(* IEC 61131-3 sources: daoli-st-library/DL_Device (part 41) *)

(* ---- FB_DL_OilLevelWatch.st ---- *)
(*
    FB_DL_OilLevelWatch —— 润滑 / 液压油油位连续监视（双阈值迟滞 + 确认延时 + NE107）
    ------------------------------------------------------------------
    组件名称  : FB_DL_OilLevelWatch
    分类      : DL_Device / LevelMonitoring
    前缀      : FB_DL_
    版本      : 1.0.0
    溯源      : 借鉴组织 —— T2-6 Rockwell AOI（矩阵行 166）：仅借鉴「设备级
                粗粒度监视 AOI」的公开功能形态（连续量监视 + 确认延时 +
                分级健康出口）；clean-room 声明 —— 零代码行复制，判据链 /
                迟滞口径 / 码位 100% 自有；非有限判据为 IEC 61131-3 标准语义
                （R79 双判）的道莅防御性实现。
    平台      : 纯 IEC 61131-3（TON / R_TRIG / LREAL 比较），CODESYS 3.5 /
                TwinCAT 3 / InoProShop / Machine Expert 通用
    作者      : 道莅代码库 · PLC编程专家（R72 构建轮 · 批 3 · 序号 9）
    ------------------------------------------------------------------
    功能说明  : 齿轮箱 / 液压单元油位巡检：欠油提前预警防干磨烧轴。
                单相监视（无顺序状态机 CASE，同族 FB_DL_AxisEncBatteryWatch
                口径家族一致）：
                ① 非有限液位闸：fLevelMm 非有限（NaN 自反判 + Inf 差值自反
                   判，R79）→ **直接故障锁存**（探头断线状态不明比欠油更
                   危险，R71 AxisEncBatteryWatch 口径家族一致），不等确认
                   延时；
                ② 组态域闸（R272 全枚举）：fLowWarnMm / fHystMm / fProbeMaxMm
                   非有限、fHystMm < 0（回差为负）、fLowWarnMm >= fProbeMaxMm
                   （阈值倒置）、fProbeMaxMm <= 0（量程非正）→ 组态锁存码
                   （根因优先归因，段 6 先于段 7）；
                ③ 双阈值迟滞判定：未预警相以进入线判（fLevelMm < fLowWarnMm），
                   已预警相以退出线判（fLevelMm >= fLowWarnMm + fHystMm），
                   防临界抖振；
                ④ TON 连续确认（断输入口径：液位回升出迟滞带 IN 即 FALSE，
                   计时清零重计）→ 预警锁存；
                ⑤ NE107 健康出口：欠油确认 → eMaintenanceReq；非有限 /
                   组态故障 → eFailure；正常 → eOk；失能 → eCheckFunction。
                锁存解除口径（R321 电平式声明）：bReset 上升沿为**唯一人工
                解除**，液位恢复越退出线为**条件恢复自动降级**双路——两路
                并存写死，禁恢复沿作唯一解除载体。预警锁存后自动降级判据 =
                液位 >= 退出线（迟滞带内保持预警，出带即自动解除）。
                满油探头饱和：fLevelMm > fProbeMaxMm → 信息级（满油合法
                工况，不拦截照判——判定方向与液位单调性一致，无危险侧偏差）。
                失能语义（R191 声明）：bEn = FALSE → bLowWarn / bError /
                nErrCode 出口清零、eHealth = eCheckFunction；_bFault /
                _bWarnLatch 锁存位**不被失能清除**（失能是操作态不是复位），
                须 bReset 上升沿解除——两语义分离。
    错误码    : 16#0003_0740 液位非有限（探头断线 / ADC 故障），直接锁存不等
                            确认延时 —— 故障级
                16#0003_0741 组态非法（阈值倒置 / 回差为负 / 阈值或量程非有限 /
                            量程非正 / 预警线不低量程上界），锁存至复位沿
                            —— 故障级
                16#0003_0742 液位越探头量程上界（探头饱和，满油合法工况）
                            —— 信息级，不置 bError（R45）
                加码反证句（R90）：0740（探头）与 0741（组态）成因互斥且调用
                方可自证（接线 vs 组态表），eHealth 出口同为 eFailure 但码位
                分流维修动作，输出组合不可互换观测，故各立一码；0742 由
                「液位在迟滞带上方 + 码位非零」唯一观测（正常满油不带码），
                不与既有输出组合重复。
    码位总账  : 16#0003_0740 用 ｜ 16#0003_0741 用 ｜ 16#0003_0742 用
    状态机    : N/A —— 单相监视，无顺序状态机，无自有 ENUM / CASE 可写；
                确认计时由 TON 实例自持（定时器状态而非顺序状态）；
                健康出口复用既有枚举 E_DL_Ne107Status（只引用）
    边界与披露: 一 TON（tonConfirm）与 R_TRIG（rtReset）每拍**无条件调用**
                   （规则 ⑦），IN 为段 7 计算出的显式条件；
                二 零全局变量、零 VAR_EXTERNAL、零物理地址；
                三 归属 Ownership：E_DL_Ne107Status 归属 I_DL_DeviceHealth.st
                   （全库唯一定义，R264），本件只引用不重声明；
                四 输入非有限 / 组态非法 → 直接锁存（不走迟滞判定集合，安全
                   侧赋值不引用本闸判定内的量，防自证循环，R127）；
                五 输出量纲：fLevelMm / fLowWarnMm / fHystMm / fProbeMaxMm 均
                   [mm]，本件不换算单位；
                六 分工互引：FB_DL_SiloLevelInterlock（料仓联锁）、
                   FB_DL_LevelSwitchVib（开关量检测）、FB_DL_HydrostaticLevelComp
                   （静压补偿换算）——本件只做模拟量油位趋势监视，不做联锁
                   与换算；
                七 依赖声明：仅 Standard.library（TON / R_TRIG / ABS），零
                   厂商方言。
    验收向量  : V1 液位 80 mm、预警线 100 mm、确认 2 s → 2 s 后 bLowWarn；
                V2 液位回升 130 mm（退出线 100 + 20）→ 自动降级解除；
                V3 液位回升 110 mm（迟滞带内）→ 预警保持（迟滞自证）；
                V4 fLevelMm = NaN → 0740 立即锁存（不等 2 s）；V5 fHystMm
                = −1 → 0741 锁存；V6 fLevelMm = 520（量程 500）→ 0742
                信息级照判；V7 bReset 上升沿 → 清锁存；V8 失能 → 出口清零、
                锁存保留。
                算法已证（脚本）：未跑 ｜ 编译器已证（三平台）：未跑
    修订记录  : 2026-11-23 v1.0.0 首次入库（R72 构建轮 · 批 3 · 序号 9）
*)
FUNCTION_BLOCK FB_DL_OilLevelWatch
VAR_INPUT
    fLevelMm    : LREAL;                   (* 油位连续值（引脚注入），[mm]，非有限即探头故障 / the oil level continuous value in mm *)
    fLowWarnMm  : LREAL := 100.0;          (* 低油位预警阈值（迟滞进入线），[mm] / the low oil warn threshold, the hysteresis enter line *)
    fHystMm     : LREAL := 20.0;           (* 迟滞回差（退出线 = 预警线 + 回差），[mm]，禁负 / the hysteresis band in mm, the exit line is warn plus band *)
    fProbeMaxMm : LREAL := 500.0;          (* 探头量程上界（饱和信息级判据），[mm]，禁非正 / the probe range upper bound in mm *)
    tConfirm    : TIME := T#2S;            (* 欠油确认延时，[ms] / the low oil confirmation delay *)
    bEn         : BOOL := TRUE;            (* 使能，[标志]，FALSE 出口清零、锁存保留 / the enable, FALSE clears the outlets, the latch kept *)
    bReset      : BOOL := FALSE;           (* 故障 / 预警复位，[标志]，上升沿唯一人工解除 / the reset, its rising edge is the only manual release *)
END_VAR
VAR_OUTPUT
    bLowWarn  : BOOL := FALSE;             (* 低油位预警锁存位（确认成立且未解除）[标志] / the low oil warn latched flag *)
    eHealth   : E_DL_Ne107Status;          (* NE107 健康出口（欠油 → eMaintenanceReq，故障 → eFailure）/ the NE 107 health outlet *)
    bValid    : BOOL := FALSE;             (* 出口可用标志，失能或锁存故障为 FALSE / the outlets usable *)
    bError    : BOOL := FALSE;             (* 故障标志，存在锁存故障时 TRUE / the fault flag *)
    nErrCode  : UDINT := 16#0000_0000;     (* 错误码，0 = 正常，锁存回放（R187）/ the error id, replayed from the latch *)
END_VAR
VAR
    _rtReset    : R_TRIG;                  (* 复位上升沿实例（无条件调用）/ the reset rising edge instance *)
    _tonConfirm : TON;                     (* 欠油确认延时实例（无条件调用）/ the low oil confirmation timer *)
    _bFault     : BOOL := FALSE;           (* 故障锁存副本（探头 / 组态），仅复位沿解除 / the internal fault latch copy *)
    _nCodeLatch : UDINT := 0;              (* 锁存成因码，故障期回放 / the latched cause code *)
    _bWarnLatch : BOOL := FALSE;           (* 预警锁存副本（自动降级或复位沿解除）/ the warn latch copy *)
    _bCfgBad    : BOOL := FALSE;           (* 组态非法标志（逐拍重算，仅用于首次锁存）/ the config fault flag *)
    _bInBad     : BOOL := FALSE;           (* 液位非有限标志（逐拍重算）/ the input fault flag *)
    _bOutDom    : BOOL := FALSE;           (* 液位越量程上界标志（逐拍重算，信息级）/ the probe saturation flag *)
    _bRun       : BOOL := FALSE;           (* 运行许可 = 使能 且 无锁存故障 / the run permit *)
    _bLowCond   : BOOL := FALSE;           (* 欠油迟滞判定条件（含自保持，送 TON）/ the low oil hysteresis condition *)
END_VAR
VAR CONSTANT
    DL_OLW_CODE_PROBE : UDINT := 16#0003_0740; (* 液位非有限锁存码 [码] / the probe fault code *)
    DL_OLW_CODE_CFG   : UDINT := 16#0003_0741; (* 组态非法锁存码 [码] / the configuration fault code *)
    DL_OLW_CODE_SAT   : UDINT := 16#0003_0742; (* 探头饱和信息码 [码] / the probe saturation info code *)
    DL_OLW_ZERO       : UDINT := 0;            (* 无符号零哨兵 [码] / the unsigned zero sentinel *)
    DL_OLW_FZERO      : LREAL := 0.0;          (* 浮点零哨兵 [mm] / the float zero sentinel *)
END_VAR

// 段 1｜出口预置（统一出口预置，R256）/ segment 1, preset every outlet
bLowWarn := FALSE;                         // 预警出口预清零（映射段回填）/ preset the warn outlet false
eHealth  := E_DL_Ne107Status.eUnknown;     // 健康出口预置未知（首拍语义）/ preset the health outlet unknown
bValid   := FALSE;                         // 可用标志预清零 / preset the usable flag false
bError   := FALSE;                         // 故障标志预清零 / preset the fault flag false
nErrCode := DL_OLW_ZERO;                   // 码位预置无错 / preset the code zero
_bLowCond := FALSE;                        // 迟滞条件预清零 / preset the condition false

// 段 2｜复位沿无条件调用（规则 ⑦）/ segment 2, the unconditional reset edge refresh
_rtReset(CLK := bReset);                   // 每拍无条件刷新 / refreshed every scan

// 段 3｜锁存解除：复位沿唯一人工解除（作用域：清双锁存 + 清码，R311 声明）/ segment 3, the manual release edge
IF _rtReset.Q THEN                         // 复位上升沿 / the reset rising edge
    _bFault := FALSE;                      // 清故障锁存（恒可达，R152 自证）/ clear the fault latch
    _bWarnLatch := FALSE;                  // 清预警锁存 / clear the warn latch
    _nCodeLatch := DL_OLW_ZERO;            // 清锁存码（可到达清除边）/ clear the latched code
END_IF

// 段 4｜组态域闸（R272 全枚举：fLowWarnMm / fHystMm / fProbeMaxMm 三引脚）/ segment 4, the configuration guard
_bCfgBad := (fLowWarnMm <> fLowWarnMm) OR ((fLowWarnMm - fLowWarnMm) <> DL_OLW_FZERO) // 预警线非有限 / the warn line non finite
         OR (fHystMm <> fHystMm) OR ((fHystMm - fHystMm) <> DL_OLW_FZERO)              // 回差非有限 / the hysteresis non finite
         OR (fProbeMaxMm <> fProbeMaxMm) OR ((fProbeMaxMm - fProbeMaxMm) <> DL_OLW_FZERO) // 量程非有限 / the range non finite
         OR (fHystMm < DL_OLW_FZERO)                                                   // 回差为负 / a negative hysteresis
         OR (fLowWarnMm >= fProbeMaxMm)                                                // 阈值倒置（预警线不低于量程上界）/ the threshold inversion
         OR (fProbeMaxMm <= DL_OLW_FZERO);                                             // 量程非正 / a non positive range

// 段 5｜输入守卫：液位非有限即危险（状态不明 > 欠油，直接锁存不等延时）/ segment 5, the input guard
_bInBad := (fLevelMm <> fLevelMm) OR ((fLevelMm - fLevelMm) <> DL_OLW_FZERO); // 液位非有限（R79 双判）/ the level non finite
_bOutDom := (fLevelMm > fProbeMaxMm);      // 液位越量程上界（探头饱和，信息级）/ the level over the range

// 段 6｜首次成因锁存（故障期内不重推断，回放锁存码，R189；组态根因优先）/ segment 6, the first cause latch
IF NOT _bFault THEN                        // 未锁存才登记 / register only while not latched
    IF _bCfgBad THEN                       // 组态非法（根因优先归因）/ the config fault first
        _bFault := TRUE;                   // 置锁存 / latch
        _nCodeLatch := DL_OLW_CODE_CFG;    // 登记组态码 / register the config code
    ELSIF _bInBad THEN                     // 液位非有限（不等确认延时）/ the probe fault, no delay
        _bFault := TRUE;                   // 置锁存 / latch
        _nCodeLatch := DL_OLW_CODE_PROBE;  // 登记探头码 / register the probe code
    END_IF
END_IF

// 段 7｜运行许可与迟滞条件（分支内不调用任何定时器）/ segment 7, the run permit and the hysteresis condition
_bRun := bEn AND (NOT _bFault);            // 使能且无锁存故障 / enabled and not latched
IF _bRun THEN                              // 运行许可成立 / the run permit holds
    IF _bWarnLatch THEN                    // 已预警相：以退出线判（迟滞防抖振）/ the latched phase, the exit line
        _bLowCond := fLevelMm < (fLowWarnMm + fHystMm); // 迟滞带内保持预警 / hold inside the band
    ELSE                                   // 未预警相：以进入线判 / the unlatched phase, the enter line
        _bLowCond := fLevelMm < fLowWarnMm; // 破进入线 / under the enter line
    END_IF
    IF _bLowCond AND _tonConfirm.Q THEN    // 破线经确认延时 / the condition confirmed
        _bWarnLatch := TRUE;               // 预警锁存 / latch the warn
    END_IF
    IF _bWarnLatch AND (NOT _bLowCond) THEN // 条件恢复自动降级（电平式双路之二，R321 声明；复位沿为人工路）/ the automatic level release
        _bWarnLatch := FALSE;              // 出迟滞带即自动解除（同拍生效）/ release over the exit line
    END_IF
ELSE                                       // 失能或锁存故障 / disabled or latched
    _bLowCond := FALSE;                    // 条件清零（TON 随之复位）/ clear the condition
END_IF

// 段 8｜确认定时器无条件调用（IN 为段 7 显式条件；断输入口径：出线即断计）/ segment 8, the unconditional confirmation timer
_tonConfirm(IN := _bRun AND _bLowCond, PT := tConfirm); // 欠油确认计时 / the confirmation timer

// 段 9｜出口映射（名实双出口同源，R191）/ segment 9, the outlet mapping
IF _bRun THEN                              // 运行许可成立 / the run permit holds
    bLowWarn := _bWarnLatch;               // 预警出口与锁存同源 / the warn outlet shares the latch
    bValid := TRUE;                        // 出口可用 / the outlets usable
    IF _bWarnLatch THEN                    // 预警确认成立 / the warn confirmed
        nErrCode := DL_OLW_ZERO;           // 预警本身不发码（欠油是正常工况分支非缺陷）/ the warn carries no code
        eHealth := E_DL_Ne107Status.eMaintenanceReq; // 欠油 → 需要维护 / maintenance required
    ELSE                                   // 无预警 / no warn
        eHealth := E_DL_Ne107Status.eOk;   // 正常 / ok
    END_IF
    IF _bOutDom AND (NOT _bWarnLatch) THEN // 运行中探头饱和且无更高优先级出口 / the saturation info
        nErrCode := DL_OLW_CODE_SAT;       // 信息级：探头饱和满油（不置 bError，R45）/ info level: the probe saturation
    END_IF
ELSIF (NOT bEn) THEN                       // 失能相（操作态优先于故障归因，同族口径）/ the disabled phase
    bLowWarn := FALSE;                     // 出口清零（锁存保留）/ the outlet cleared, the latch kept
    bError := FALSE;                       // 失能不是故障 / a disabled block is not a fault
    nErrCode := DL_OLW_ZERO;               // 失能不发码 / no code while disabled
    eHealth := E_DL_Ne107Status.eCheckFunction; // 失能 → 功能检查 / function check
ELSE                                       // 锁存故障相（失能优先级之上）/ the latched fault phase
    bLowWarn := FALSE;                     // 故障相预警出口清零（归并故障出口）/ the warn outlet cleared
    bError := TRUE;                        // 故障标志置位 / raise the fault flag
    nErrCode := _nCodeLatch;               // 回放锁存码 / replay the latched code
    eHealth := E_DL_Ne107Status.eFailure;  // 故障 → 失效（信号不可信）/ failure
END_IF
END_FUNCTION_BLOCK

(* ---- FB_DL_PressureReliefMonitor.st ---- *)
(*==============================================================================
 * 组件名称 (Component)  : FB_DL_PressureReliefMonitor
 * 溯源说明 (Provenance): 道莅 clean-room 防御性实现（IEC 61131-3 纯净实现，闭源文档仅借语义，零代码行）
 * 所属子库 (Sublibrary) : DL_Device / SafetyMonitor
 * 当前版本 (Version)    : 1.0.0
 * 兼容性   (Platform)   : CODESYS 3.5 / TwinCAT 3 / 汇川 InoProShop / 施耐德
 *                         Machine Expert；纯 IEC 61131-3（第 3 版），仅用
 *                         Standard.library 的 TON / ABS / MAX
 * 组件分类 (Category)   : 功能块（FUNCTION_BLOCK）· 安全阀起跳/回座监视与台账
 * 功能一句话 (Summary)  : 用阀前/阀后压力判安全阀是否起跳，累计动作次数与累计
 *                         开启时长，给出本次起跳峰值压力与 NE107 健康分级。
 *
 * 本件存在的意义 (Why this unit exists)
 *   过程安全台账要求「安全阀一年动作了几次、累计开启多久」——这是法检项。
 *   库内 AlarmManager 数的是报警不是阀门动作，PortDiag 系列数的是通讯事件，
 *   没有任何件维护这张台账。同时「阀前持续超整定而阀后不同步升高」是
 *   安全阀不泄放的典型特征，属于必须报出来的失效形态。
 *
 * 台账纪律 (Ledger discipline)
 *   ① 起跳判据必须用**回座比做迟滞**（fUpPressure < fSetPressure × fBlowdown），
 *      硬阈值会让压力在整定点附近抖动并反复计数——这是台账失真的头号原因；
 *   ② 单次起跳时长 < tMinLift 不计入 nLiftCount（信息 0175）：工艺压力波动
 *      引起的瞬时顶开不构成「动作」，但仍计入累计开启时长之外的判定之外，
 *      两者口径不同，头注释写死；
 *   ③ 计数与累计时长累加前判上界，饱和不回绕（R35）；TIME 溢出用比较式
 *      预判（R54），比较表达式内不出现加乘运算符；
 *   ④ **失能不清台账**：计数、累计时长、峰值一律保持；若失能发生在起跳期间，
 *      以失能拍作为该次起跳的结束拍如实入账，绝不丢一次真实动作。
 *
 * 健康映射（写死在此，不散落实现体）
 *   参数非法 / 输入非有限                        → eFailure
 *   起跳中且阀后压力 > 整定 × DL_DN_FAIL_RATIO    → eFailure（疑似不泄放）
 *   nLiftCount >= uMaintLimit                    → eMaintenanceReq
 *   其余（有判定能力）                            → eOk
 *   未使能（无判定能力）                          → eUnknown
 *   DL_DN_FAIL_RATIO = 0.5 为件内经验阈值：安全阀正常起跳时阀后应接近大气，
 *   若阀后压力仍高于整定的一半，说明介质没有真正排出去（下游堵塞或阀瓣卡滞）。
 *
 * 边界安全 (Boundary)
 *   - fSetPressure <= 0 或 fBlowdown 不在 (0, 1) 或非有限 → 故障 033F、bValid = FALSE，
 *     **台账保持不动**（参数错了不等于阀门没动作过）；
 *   - 任一压力非有限 → 故障 0340，**保持 bLifted 与计数不变**（坏值不得伪造动作）；
 *   - bError 的每一个置位源都能在 eErr 找到对应码（R45 纪律）；
 *   - CASE 落 ELSE 置 0341 兜底并回 eFault；
 *   - 本件无复位引脚：台账只能靠 FB 实例重建清零（法检台账不允许被误复位，
 *     这是刻意设计，已留档）。
 *
 * 错误码    : 16#0003_0174 起跳事件已记录（动作次数 +1，累计时长继续累加）——信息级
 *             16#0003_0175 单次起跳时长低于 tMinLift，按工艺波动滤除不计入台账——信息级
 *             16#0003_033F 整定压力或回座比非法——故障级，bValid = FALSE
 *             16#0003_0340 压力输入非有限，保持台账与判定不变——故障级，坏值不得伪造动作
 *             16#0003_0341 状态机落 ELSE 兜底（非法状态）——故障级，回 eIdle 并保持台账
 * 码位总账  : 16#0003_0174 用 / 16#0003_0175 用 ｜ 16#0003_033F 用 / 16#0003_0340 用 / 16#0003_0341 用
 * 状态机    : E_DL_ReliefState（eIdle / eLifted / eReseat / eFault），CASE 含 ELSE 兜底，
 *             ELSE 置 16#0003_0341 并回 eFault；失能回 eIdle 但台账保持
 * 采样约定  : 每任务周期调用一次；时长按滚动时钟差累加（上拍快照，R45②）
 * 依赖说明  : 仅 Standard.library；健康出口引用 E_DL_Ne107Status（属主 I_DL_DeviceHealth，
 *             **引用不重声明**，R70③）
 * 验收向量  : V1 压力从 8 缓升到 10.5 bar 持续 200 ms → eLifted，bLifted = TRUE，
 *                fPeakPressure 跟随峰值；压力回落到 8.9（< 10×0.90 = 9.0）→ eReseat，
 *                时长 ≥ 500 ms 时 nLiftCount + 1 且 eErr = 0174，eHealth 随计数升级
 *             V2 起跳仅 300 ms（< tMinLift 500 ms）→ nLiftCount 不变，eErr = 0175（滤除主向量）
 *             V3 起跳中阀后压力 6 bar（> 10×0.5）→ eHealth = eFailure（不泄放主向量）
 *             V4 fBlowdown = 1.2 → 033F，bValid = FALSE，nLiftCount 与 tOpenTotal 保持
 *             V5 fUpPressure = NaN → 0340，bLifted 与计数保持（坏值不伪造动作主向量）
 *             V6 压力在 9.98~10.02 之间抖动 → 不重复计数（回座迟滞主向量）
 *             V7 bEnable 落于起跳中 → eIdle，本次时长如实入账，计数不清零
 * 红线自检  : 全局变量声明零使用 / 外部变量访问零使用 / 物理地址零使用 ｜ 纯 IEC 61131-3 ｜ 无除法
 *             浮点只用大小与容差比较 ｜ 无循环 ｜ 全变量双语同行注释 ｜ ENUM + CASE
 *             含 ELSE ｜ TON 在主体前部无条件刷新 ｜ TIME 溢出比较式预判 ｜
 *             阈值常量化，无魔法数
 * 修订历史  : 2026-11-16  v1.0.0  首版入库（R22 · 批 2 · 设备安全台账）
 *============================================================================*)

(*-----------------------------------------------------------------------------
 * 枚举: E_DL_ReliefState（归属本功能块，同文件发布，全库唯一定义）
 * 含义: 安全阀监视的工作相位。0 起步长 10。
 * 注意: 健康出口类型 E_DL_Ne107Status 属主为 I_DL_DeviceHealth（DL_Device 契约件），
 *       本件只引用、不重声明（R70③ 全库唯一定义）。
 *-----------------------------------------------------------------------------*)
TYPE E_DL_ReliefState :
(
    eIdle   := 0,      // 待机：未起跳，等待起跳确认 / Idle, waiting for a confirmed lift
    eLifted := 10,     // 起跳中：阀前高于整定，正在累计时长 / Lifted, upstream above the set pressure
    eReseat := 20,     // 回座：单拍入账相，随后回待机 / Reseat, one scan to book the event
    eFault  := 99      // 故障：参数非法或输入非有限 / Fault, illegal parameter or non-finite input
);
END_TYPE

FUNCTION_BLOCK FB_DL_PressureReliefMonitor
VAR_INPUT
    fUpPressure  : REAL;                       // 阀前压力 [bar g] / upstream pressure [bar g]
    fDnPressure  : REAL;                       // 阀后压力 [bar g] / downstream pressure [bar g]
    fSetPressure : REAL := 10.0;               // 整定压力 [bar g]，须 > 0 / set pressure [bar g], must be > 0
    fBlowdown    : REAL := 0.90;               // 回座压力比 [倍]，须在 0~1 之间 / reseat ratio [ratio], must lie inside zero and one
    tConfirm     : TIME := T#200MS;            // 起跳确认时间 [ms] / lift confirm time [ms]
    tMinLift     : TIME := T#500MS;            // 最短起跳时长 [ms]，低于此按波动滤除 / minimum lift duration [ms], shorter ones are filtered
    uMaintLimit  : UINT := 50;                 // 动作次数维护门限 [次] / maintenance count threshold [count]
    bEnable      : BOOL;                       // 使能（失能不清台账） / enable, the ledger survives a disable
END_VAR
VAR_OUTPUT
    bLifted      : BOOL;                       // 当前处于起跳状态 / currently lifted
    nLiftCount   : UDINT;                      // 累计动作次数 [次] / accumulated lift count [count]
    tOpenTotal   : TIME;                       // 累计开启时长 [ms] / accumulated open time [ms]
    fPeakPressure : REAL;                      // 本次起跳峰值压力 [bar g] / peak upstream pressure of the current lift [bar g]
    eHealth      : E_DL_Ne107Status;           // NE107 健康分级（引用唯一属主） / NE107 health status, referenced from its owner
    eErr         : UDINT;                      // 错误码，0 表示无错 / error code, 0 means no error
    bError       : BOOL;                       // 故障级标志，仅故障级错误置位 / fault-class flag, set only on fault-level codes
    bValid       : BOOL;                       // 输出可用标志 / outputs usable flag
END_VAR
VAR
    fbConfirm    : TON;                        // 起跳确认计时，段 5 无条件刷新 [ms] / lift confirm timer
    fbElapsed    : TON;                        // 滚动时钟，段 5 无条件刷新 [ms] / rolling elapsed clock
    _eState      : E_DL_ReliefState := E_DL_ReliefState.eIdle; // 当前相位 / current phase
    _bInit       : BOOL := FALSE;              // 首扫标志，初值 FALSE 取非判定 / first-scan flag, tested negated
    _bParamBad   : BOOL;                       // 参数非法标志 / illegal parameter flag
    _bFiniteBad  : BOOL;                       // 输入非有限标志 / non-finite input flag
    _bIllegal    : BOOL;                       // 非法状态标志 / illegal state flag
    _bAbove      : BOOL;                       // 阀前高于整定（确认条件） / upstream above the set pressure
    _bReseatNow  : BOOL;                       // 回座判据成立 / reseat criterion satisfied
    _bConfBreak  : BOOL;                       // 确认计时器断输入一拍 / confirm timer one-scan break
    _bElapsedBreak : BOOL;                     // 滚动时钟断输入一拍 / rolling clock one-scan break
    _bNoRelief   : BOOL;                       // 疑似不泄放标志 / suspected no-relief flag
    _bBooked     : BOOL;                       // 本拍已入账标志 / booked this scan flag
    _bReseatPulse : BOOL;                      // 回座单拍脉冲（入账触发） / reseat one-scan pulse, triggers the booking
    _bLiftedPrev : BOOL;                       // 本拍进入时的起跳相快照（R38 镜像量） / lifted snapshot taken before the transitions
    _tConfirmUse : TIME := T#200MS;            // 生效确认时间 [ms]，已钳位 / effective confirm time, clamped
    _tMinLiftUse : TIME := T#500MS;            // 生效最短起跳时长 [ms]，已钳位 / effective minimum lift, clamped
    _tEtPrev     : TIME;                       // 滚动时钟上拍快照 [ms] / previous scan snapshot of the clock
    _tDelta      : TIME;                       // 本拍时长增量 [ms] / elapsed increment of this scan
    _tLiftDur    : TIME;                       // 本次起跳已持续时长 [ms] / duration of the current lift [ms]
    _tTotalAcc   : TIME;                       // 累计开启时长保持量 [ms] / held accumulated open time [ms]
    _uCountAcc   : UDINT;                      // 累计动作次数保持量 [次] / held lift count [count]
    _fPeakAcc    : REAL;                       // 本次起跳峰值保持量 [bar g] / held peak pressure of the current lift [bar g]
    _fPeakTot    : REAL;                       // 历史峰值（供 HMI 参考） [bar g] / historical peak pressure [bar g]
END_VAR
VAR CONSTANT
    DL_VAL_LIM   : REAL := 1.0E6;              // 有限性判定的绝对值上限 [bar g] / finiteness ceiling [bar g]
    DL_SET_MIN   : REAL := 0.0;                // 整定压力下限 [bar g]，须严格大于 / set pressure floor, strictly greater
    DL_BLOW_MIN  : REAL := 0.0;                // 回座比下限 [倍]，须严格大于 / reseat ratio floor, strictly greater
    DL_BLOW_MAX  : REAL := 1.0;                // 回座比上限 [倍]，须严格小于 / reseat ratio ceiling, strictly less
    DL_DN_FAIL_RATIO : REAL := 0.5;            // 阀后不泄放判据比 [倍]，件内经验阈值 / no-relief ratio, an empirical in-unit threshold
    DL_CONF_MAX_MS : DINT := 60000;            // 确认时间上限 [ms] / confirm time ceiling [ms]
    DL_MINLIFT_MAX_MS : DINT := 3600000;       // 最短起跳时长上限 [ms]，一小时 / minimum lift ceiling, one hour
    DL_TIME_ZERO : TIME := T#0MS;              // 时间零值基准 [ms] / time zero reference
    DL_ROLL      : TIME := T#1H;               // 滚动时钟周期 [ms]，到顶重启防 ET 停滞 / rolling clock period, restarted at the top
    DL_TOTAL_MAX : TIME := T#24H;              // 累计时长饱和上界 [ms] 上限值：判溢出用 / accumulation ceiling, used by the overflow test
    DL_TIME_SAT  : TIME := T#24H;              // 累计时长饱和输出值 [ms] / accumulation saturation value
    DL_CNT_MAX   : UDINT := 16#FFFF_FFFF;      // 计数饱和上界 [次]，不回绕 / counter saturation ceiling, never wraps
END_VAR

(*------------------------------------------------------------------------------
 * 段 1｜每拍预置（台账保持量不预置；输出在段 9 单点写入）
 *      Per-scan presets, the ledger values are never cleared here
 *-----------------------------------------------------------------------------*)
eErr         := 16#0000_0000;                  // 错误码每拍重算 / error code recomputed every scan
bError       := FALSE;                         // 故障标志每拍重算 / fault flag recomputed every scan
bValid       := FALSE;                         // 可用标志每拍重算 / usable flag recomputed every scan
_bParamBad   := FALSE;                         // 参数非法标志预清零 / parameter flag pre-cleared
_bFiniteBad  := FALSE;                         // 非有限标志预清零 / non-finite flag pre-cleared
_bIllegal    := FALSE;                         // 非法状态标志预清零 / illegal state flag pre-cleared
_bAbove      := FALSE;                         // 超整定条件预置 FALSE / above-set condition preset FALSE
_bReseatNow  := FALSE;                         // 回座判据预置 FALSE / reseat criterion preset FALSE
_bNoRelief   := FALSE;                         // 不泄放标志预置 FALSE / no-relief preset FALSE
_bBooked     := FALSE;                         // 入账标志预置 FALSE / booked flag preset FALSE
_bReseatPulse := FALSE;                        // 回座脉冲预置 FALSE / reseat pulse preset FALSE
_bLiftedPrev := FALSE;                         // 起跳快照预置 FALSE / lifted snapshot preset FALSE

(*------------------------------------------------------------------------------
 * 段 2｜首扫初始化（台账全部从零起，峰值从当前阀前压力起）
 *      First-scan initialisation, the ledger starts at zero
 *-----------------------------------------------------------------------------*)
IF NOT _bInit THEN
    _eState     := E_DL_ReliefState.eIdle;     // 相位待机 / phase idle
    _uCountAcc  := 0;                          // 动作次数清零 [次] / lift count cleared
    _tTotalAcc  := DL_TIME_ZERO;               // 累计时长清零 [ms] / accumulated time cleared
    _tLiftDur   := DL_TIME_ZERO;               // 本次时长清零 [ms] / current lift duration cleared
    _tEtPrev    := DL_TIME_ZERO;               // 时钟快照清零 [ms] / clock snapshot cleared
    _fPeakAcc   := 0.0;                        // 本次峰值清零 [bar g] / current peak cleared
    _fPeakTot   := 0.0;                        // 历史峰值清零 [bar g] / historical peak cleared
    _bConfBreak := TRUE;                       // 确认计时从零开始 / confirm timer starts from zero
    _bElapsedBreak := TRUE;                    // 滚动时钟从零开始 / rolling clock starts from zero
    _bInit      := TRUE;                       // 首扫只做一次 / the first scan runs once
END_IF

(*------------------------------------------------------------------------------
 * 段 3｜参数闸门（整定压力与回座比；非法只降可用性，台账一律保持）
 *      Parameter gate, an illegal parameter lowers usability but never touches the ledger
 *-----------------------------------------------------------------------------*)
IF (fSetPressure <> fSetPressure) OR (ABS(fSetPressure) > DL_VAL_LIM) OR (fSetPressure <= DL_SET_MIN) THEN
    _bParamBad := TRUE;                        // 整定压力非法 / set pressure illegal
END_IF
IF (fBlowdown <> fBlowdown) OR (fBlowdown <= DL_BLOW_MIN) OR (fBlowdown >= DL_BLOW_MAX) THEN
    _bParamBad := TRUE;                        // 回座比非法（须严格在 0~1 之间） / reseat ratio illegal
END_IF

(*------------------------------------------------------------------------------
 * 段 4｜压力输入有限性（区间判据同时拦 NaN 与 ±Inf）
 *      Pressure finiteness, the interval test catches NaN and infinity
 *-----------------------------------------------------------------------------*)
IF (fUpPressure < -DL_VAL_LIM) OR (fUpPressure > DL_VAL_LIM) THEN
    _bFiniteBad := TRUE;                       // 阀前压力非有限 / upstream pressure non-finite
END_IF
IF (fDnPressure < -DL_VAL_LIM) OR (fDnPressure > DL_VAL_LIM) THEN
    _bFiniteBad := TRUE;                       // 阀后压力非有限 / downstream pressure non-finite
END_IF

(*------------------------------------------------------------------------------
 * 段 5｜计时器无条件刷新（R40）+ 本拍时长增量（R45② 上拍快照）
 *      Timers refreshed unconditionally, the elapsed increment uses a previous-scan snapshot
 *-----------------------------------------------------------------------------*)
_tConfirmUse := tConfirm;                      // 确认时间直取引脚 [ms] / confirm time from the pin
IF TIME_TO_DINT(_tConfirmUse) > DL_CONF_MAX_MS THEN
    _tConfirmUse := DINT_TO_TIME(DL_CONF_MAX_MS); // 超上限钳位（无专用码位，R90 不新开码） / clamped
END_IF
IF TIME_TO_DINT(_tConfirmUse) < 0 THEN
    _tConfirmUse := DL_TIME_ZERO;              // 负时间结构性不可达，兜底为 0 / structurally unreachable fallback
END_IF

_tMinLiftUse := tMinLift;                      // 最短起跳时长直取引脚 [ms] / minimum lift from the pin
IF TIME_TO_DINT(_tMinLiftUse) > DL_MINLIFT_MAX_MS THEN
    _tMinLiftUse := DINT_TO_TIME(DL_MINLIFT_MAX_MS); // 超上限钳位 / clamped
END_IF
IF TIME_TO_DINT(_tMinLiftUse) < 0 THEN
    _tMinLiftUse := DL_TIME_ZERO;              // 负时间兜底为 0 / fallback to zero
END_IF

IF NOT _bFiniteBad THEN
    _bAbove := (fUpPressure > fSetPressure);   // 超整定判据 [布尔] / above-set test
    IF NOT _bParamBad THEN
        _bReseatNow := (fUpPressure < (fSetPressure * fBlowdown)); // 回座判据：低于整定×回座比 / reseat test
    END_IF
    _bNoRelief := (fDnPressure > (fSetPressure * DL_DN_FAIL_RATIO)); // 阀后未降：疑似不泄放 / downstream not relieved
END_IF

fbConfirm(IN := _bAbove AND (NOT _bConfBreak), PT := _tConfirmUse); // 起跳确认计时
_bConfBreak := FALSE;                          // 断输入拍在调用后自清 / break self-cleared after the call

fbElapsed(IN := (NOT _bElapsedBreak), PT := DL_ROLL); // 滚动时钟无条件刷新
_bElapsedBreak := FALSE;                       // 断输入拍在调用后自清 / break self-cleared
_tDelta := fbElapsed.ET - _tEtPrev;            // 本拍增量 = 当前 ET − 上拍快照 / increment from the snapshot
IF TIME_TO_DINT(_tDelta) < 0 THEN
    _tDelta := DL_TIME_ZERO;                   // 时钟重启拍：增量按 0 处理，绝不倒扣 / restart scan counts as zero
END_IF
_tEtPrev := fbElapsed.ET;                      // 快照在本拍末更新（唯一写入点） / snapshot updated once
IF fbElapsed.Q THEN
    _bElapsedBreak := TRUE;                    // 到顶重启：下一拍 ET 归零 / restart so the next scan starts from zero
    _tEtPrev := DL_TIME_ZERO;                  // 重启后快照同步归零 / the snapshot follows the restart
END_IF

(* 起跳相快照在迁移之前采集（R38）：迁移拍也要把本拍时长增量算进本次起跳 *)
(* The lifted snapshot is taken before the transitions so the final scan still counts *)
_bLiftedPrev := (_eState = E_DL_ReliefState.eLifted);

(*------------------------------------------------------------------------------
 * 段 6｜相位机（只做迁移；台账入账在段 7，出口在段 9）
 *      Phase machine, transitions only, the ledger is booked in segment seven
 *-----------------------------------------------------------------------------*)
CASE _eState OF

    E_DL_ReliefState.eIdle:                    // 待机：确认超整定即起跳
        IF _bParamBad OR _bFiniteBad THEN
            _eState := E_DL_ReliefState.eFault; // 原因未消失，转故障 / the cause persists
        ELSIF bEnable AND fbConfirm.Q THEN
            _eState     := E_DL_ReliefState.eLifted; // 进起跳相 / enter the lifted phase
            _tLiftDur   := DL_TIME_ZERO;       // 本次时长从零累计 / duration starts at zero
            _fPeakAcc   := fUpPressure;        // 峰值初值 = 起跳压力 / the peak starts at the lift pressure
            _bNoRelief  := FALSE;              // 起跳首拍不判不泄放 / no no-relief verdict on the first scan
        ELSIF NOT bEnable THEN
            _eState := E_DL_ReliefState.eIdle; // 失能保持待机，台账不动 / disabled, the ledger is untouched
        END_IF

    E_DL_ReliefState.eLifted:                  // 起跳中：回座或失能都结束本次起跳
        IF _bFiniteBad THEN
            _eState := E_DL_ReliefState.eFault; // 坏值：保持判定与台账（段 7 不入账） / non-finite, hold everything
        ELSIF _bParamBad THEN
            _eState := E_DL_ReliefState.eFault; // 参数非法：转故障 / illegal parameters go to fault
        ELSIF NOT bEnable THEN
            _eState := E_DL_ReliefState.eReseat; // 失能以本拍作为结束拍，如实入账 / disabling closes the lift honestly
        ELSIF _bReseatNow THEN
            _eState := E_DL_ReliefState.eReseat; // 回座 / reseated
        END_IF

    E_DL_ReliefState.eReseat:                  // 回座：单拍入账相（**本相不在此迁移**，先入账后迁移）
        _bReseatPulse := TRUE;                 // 置入账脉冲，迁移交给段 7 入账之后 / book first, transition after

    E_DL_ReliefState.eFault:                   // 故障：参数合法且输入有限才回待机
        IF bEnable AND (NOT _bParamBad) AND (NOT _bFiniteBad) THEN
            _eState := E_DL_ReliefState.eIdle; // 原因消失，回待机并重新确认 / cause cleared, confirm again
            _bConfBreak := TRUE;               // 确认计时重启，避免沿用故障期残留 / restart the confirm timer
        END_IF

    ELSE
        _bIllegal := TRUE;                     // 标记非法状态 / flag the illegal state
        _eState   := E_DL_ReliefState.eFault;  // 回故障态 / back to the fault state
        eErr      := 16#0003_0341;             // 故障级：状态机兜底 / fault: state machine fallback
        bError    := TRUE;                     // 置故障标志 / raise the fault flag
END_CASE

(*------------------------------------------------------------------------------
 * 段 7｜台账演进（唯一累加点：起跳相按时长增量，回座相一次性入账）
 *      Ledger evolution, the single accumulation point
 *-----------------------------------------------------------------------------*)
IF _bLiftedPrev AND (NOT _bFiniteBad) AND (NOT _bParamBad) THEN
    _tLiftDur := _tLiftDur + _tDelta;          // 本次起跳时长累加 [ms] / current lift duration accumulates
    IF fUpPressure > _fPeakAcc THEN
        _fPeakAcc := fUpPressure;              // 跟踪本次峰值 [bar g] / track the current peak
    END_IF
    IF fUpPressure > _fPeakTot THEN
        _fPeakTot := fUpPressure;              // 跟踪历史峰值 [bar g] / track the historical peak
    END_IF
    IF _tTotalAcc > (DL_TOTAL_MAX - _tDelta) THEN
        _tTotalAcc := DL_TIME_SAT;             // 饱和不回绕（R54 比较式预判） [ms] / saturate, never wrap
    ELSE
        _tTotalAcc := _tTotalAcc + _tDelta;    // 累计开启时长 [ms] / accumulate the open time
    END_IF
END_IF

(* 回座（或失能结束起跳）的当拍一次性入账，入账之后再迁移回待机 *)
(* Book the event once on the reseat scan, then transition back to idle *)
IF _bReseatPulse AND (NOT _bBooked) THEN
    _bBooked := TRUE;                          // 本拍只入账一次 / book exactly once
    IF TIME_TO_DINT(_tLiftDur) >= TIME_TO_DINT(_tMinLiftUse) THEN
        IF _uCountAcc < DL_CNT_MAX THEN
            _uCountAcc := _uCountAcc + 1;      // 动作次数 +1（饱和不回绕） [次] / count incremented
        END_IF
        eErr := 16#0003_0174;                  // 信息级：起跳事件已记录 / informational: lift event recorded
    ELSE
        eErr := 16#0003_0175;                  // 信息级：时长不足，按工艺波动滤除 / informational: filtered as process fluctuation
    END_IF
    _tLiftDur := DL_TIME_ZERO;                 // 本次时长清零，准备下一次 / reset the duration
END_IF

(* 入账完成后才允许迁移：次序不可反（先入账、后迁移，R45） *)
(* Transition only after the booking, the order cannot be reversed *)
IF _eState = E_DL_ReliefState.eReseat THEN
    _eState := E_DL_ReliefState.eIdle;         // 回待机，重新等待起跳确认 / back to idle and wait for the next confirm
END_IF

(*------------------------------------------------------------------------------
 * 段 8｜故障码单一优先级链（每一个 bError 置位源都在此找到对应码，R45）
 *      Single priority chain of fault codes, every bError source maps to a code
 *-----------------------------------------------------------------------------*)
IF _bIllegal THEN
    bError := TRUE;                            // 非法状态已置码 0341（CASE 兜底） / illegal state, code 0341 set by the fallback
ELSIF _bParamBad THEN
    eErr   := 16#0003_033F;                    // 故障级：整定压力或回座比非法 / fault: set pressure or reseat ratio illegal
    bError := TRUE;                            // 置故障标志 / raise the fault flag
ELSIF _bFiniteBad THEN
    eErr   := 16#0003_0340;                    // 故障级：压力输入非有限，台账保持 / fault: non-finite pressure, ledger held
    bError := TRUE;                            // 置故障标志 / raise the fault flag
END_IF

(*------------------------------------------------------------------------------
 * 段 9｜健康分级（等级→健康映射集中在此，不散落实现体）
 *      Health grading, the whole mapping lives here
 *-----------------------------------------------------------------------------*)
IF _bParamBad OR _bFiniteBad OR _bIllegal THEN
    eHealth := E_DL_Ne107Status.eFailure;      // 参数非法或输入非有限：失效 / illegal parameter or non-finite input
ELSIF (_eState = E_DL_ReliefState.eLifted) AND _bNoRelief THEN
    eHealth := E_DL_Ne107Status.eFailure;      // 起跳中阀后未降：疑似不泄放 / lifted but downstream not relieved
ELSIF _uCountAcc >= uMaintLimit THEN
    eHealth := E_DL_Ne107Status.eMaintenanceReq; // 动作次数达门限：需维护 / maintenance threshold reached
ELSIF NOT bEnable THEN
    eHealth := E_DL_Ne107Status.eUnknown;      // 未使能：无判定能力 / no verdict capability while disabled
ELSE
    eHealth := E_DL_Ne107Status.eOk;           // 其余：正常 / otherwise normal
END_IF

(*------------------------------------------------------------------------------
 * 段 10｜出口单点写入与可用性仲裁
 *      Single write point of the outputs and the usability arbitration
 *-----------------------------------------------------------------------------*)
bLifted       := (_eState = E_DL_ReliefState.eLifted); // 起跳状态出口 / lifted outlet
nLiftCount    := _uCountAcc;                   // 动作次数出口 [次] / lift count outlet
tOpenTotal    := _tTotalAcc;                   // 累计开启时长出口 [ms] / accumulated open time outlet
fPeakPressure := _fPeakAcc;                    // 本次起跳峰值出口 [bar g] / current lift peak outlet

IF bError THEN
    bValid := FALSE;                           // 故障级：输出不可用（台账仍如实上报） / fault: unusable, the ledger is still reported
ELSIF NOT bEnable THEN
    bValid := FALSE;                           // 失能：判定不可用（台账保持） / disabled: no verdict, ledger held
ELSIF _bFiniteBad THEN
    bValid := FALSE;                           // 非有限拍：判定不可用 / non-finite scan: no verdict
ELSE
    bValid := TRUE;                            // 判定可用 / verdict usable
END_IF

END_FUNCTION_BLOCK

(* ---- FB_DL_PulseDirStepper.st ---- *)
(*==============================================================================
 * 组件名称 (Component)  : FB_DL_PulseDirStepper
 * 所属子库 (Sublibrary) : DL_Device
 * 当前版本 (Version)    : 1.0.1
 * 分类     (Category)   : 设备功能块（Function Block · 脉冲方向型开环步进控制器）
 * 作者     (Author)     : Daoli Library
 * 日期     (Date)       : 2026-11-15
 * 兼容性   (Platform)   : CODESYS 3.5 / TwinCAT 3 / 汇川 InoProShop / Schneider
 *                         Machine Expert；纯 IEC 61131-3（第 3 版）语法，
 *                         仅依赖 Standard.library（TON），零厂商方言
 * 功能简介 (Function)   : 脉冲 + 方向型开环步进控制器，实现接口
 *                         I_DL_StepperOpenLoop 的全部属性与方法。① 梯形加减速
 *                         脉冲频率规划（加速/匀速/减速三段，短行程退化为三角型）；
 *                         ② 限位保护（同向限位立即停发脉冲并锁故障，方向拒绝为
 *                         电平判据持续生效）；③ 堵转超时判据（运动耗时超理论耗时
 *                         乘裕度系数加附加裕度即判故障）；④ 脉冲按任务周期定宽
 *                         输出（R24：脉宽恒为一拍，停发在本拍内完成，无半脉冲）。
 * 职责边界 (Scope)      : 不绑定输出模块（脉冲/方向/使能全部经引脚输出，物理口
 *                         映射由适配层完成）；不做位置闭环（开环无编码器，位置为
 *                         指令推算值）；不做回原与点动（由上层组合实现）；不构成
 *                         ISO 13849 / IEC 62061 认证安全功能，急停与安全门必须由
 *                         认证安全回路在输出侧直接切断。
 * 开源溯源 (Origin)     : 来源标签 stepper（GitHub topics 开组）+ plcopen-motion
 *                         梯形规划语义。仅参考 MIT 许可开源步进驱动项目（AccelStepper
 *                         及同类公开仓库）公开的「梯形加减速脉冲频率规划算法思想」
 *                         与「脉冲当量 / 最大速度 / 加速度 / 超时」参数域惯例，以及
 *                         PLCopen 公开规范中梯形速度曲线的段划分语义；枚举编号、
 *                         状态机、限位/堵转判据、故障码位与脉冲发生实现 100% 本库
 *                         独立设计，clean-room 实现，未复制任何来源代码行，不构成
 *                         任何来源的衍生作品。
 * 公约遵循 (Convention) : 0.1/R19 首扫范式；0.2/R21 bError 排除信息级码；0.5/R7
 *                         定时器实例主体最前部无条件刷新；0.6/R14 定时器语义参数
 *                         变化断输入一拍；0.7/R15 故障锁存仅复位路径清码；0.9 非
 *                         有限值防御与出口默认值先赋；0.12/R22 接口属性以 PROPERTY
 *                         GET 承载、非接口成员保留引脚；0.14 除法防零与浮点容差；
 *                         0.15 单位统一 mm / mm/s / mm/s² / Hz / 脉冲；0.16 全常量化。
 * 红线自检 (Redline)    : 全局隔离 ✓｜命名合规 ✓｜注释完整 ✓（声明行全中英双语）｜
 *                         OOP 封装 ✓（IMPLEMENTS 接口、状态私有、属性只读）｜周期
 *                         安全 ✓（TON 无条件刷新，方法无跨周期驻留）｜防御编程 ✓
 *                         （除零守卫、浮点容差、CASE+ELSE 兜底、脉宽下限保护）｜
 *                         可移植性 ✓（纯 IEC 61131-3）｜终结符成对 ✓
 * 设计要点 (Key notes)  : ① 频率上限硬约束：脉冲每拍最多翻转一次，最高频率为
 *                         1 / (2 × 任务周期)（一高拍 + 一低拍）；超限即钳位并置
 *                         0003_0131，保证脉宽下限恒为一拍（R24）。
 *                         ② 梯形解析式（脉冲域，速度为频率）：加速段步数 na =
 *                         v² / (2a)；若 2 × na > N 则三角型，na = N / 2 且峰值
 *                         v = SQRT(a × N)；理论耗时 t = 2(v/a) + (N − 2na)/v [s]。
 *                         ③ 堵转判据：时限 = t × 1.5 + tStallTimeout，定时器自运动
 *                         起点计时，到期判堵转（开环无反馈，只能以时间偏离推断）。
 *                         ④ 限位语义：运动中同向限位即停发并锁故障；复位后方向拒绝
 *                         仍由开关电平承担（停在限位开关上时仅反方向可动），避免
 *                         「卡在限位无法脱离」的死锁。
 *                         ⑤ 故障不切使能：bEnableOut 恒透传使能指令，故障期保持保持
 *                         力矩，防垂直轴溜车；切使能由上层安全回路决定。
 * 偏离留档 (Deviation)  : ① 规格 OUT 列的 bReady / fPosition / uAlarmWord 标为
 *                         「接口属性实现」，按公约 0.12 改为 PROPERTY GET 承载
 *                         （读法不变，语义一致）；② 规格 VAR 段 bFirstScan 改名
 *                         _bInit（公约 0.1）；③ 规格建议故障码 0003_0230~0235 与
 *                         既有 FB_DL_VacuumEjector（0230~0232）冲突，依公约 0.8
 *                         顺延至 0003_02E0~02E4；信息级扩至 0136。
 * 故障码表 (Error codes) :
 *                         16#0003_0130【信息级】速度指令超最大速度已钳位
 *                         16#0003_0131【信息级】脉冲频率超任务周期上限已钳位
 *                         16#0003_0132【信息级】位移不足一个脉冲当量被忽略
 *                         16#0003_0133【信息级】运动/复位指令被拒绝（状态不满足）
 *                         16#0003_0134【信息级】限位方向禁止（同向指令被拒）
 *                         16#0003_0135【信息级】去使能冻结脉冲输出
 *                         16#0003_0136【信息级】任务周期非法已兜底为 10 ms
 *                         16#0003_0137【信息级】减速收尾残差不足一脉冲，按到位处理
 *                         16#0003_02E0【故障级】组态参数非法（Init 参数域越界）
 *                         16#0003_02E1【故障级】限位入侵停机（运动中同向限位触发）
 *                         16#0003_02E2【故障级】驱动器报警输入有效
 *                         16#0003_02E3【故障级】堵转超时（超理论耗时乘裕度）
 *                         16#0003_02E4【故障级】非法状态兜底（枚举越界）
 * 验收向量 (Acceptance) :
 *   V1 规划：当量 400、细分 1、速度 20 mm/s、加速度 500 mm/s²、行程 10 mm →
 *      总步数 4000、指令频率 8000 Hz（必被钳位）、加速段按 v²/(2a) 复算一致；
 *   V2 钳位：任务周期 10 ms → 上限 50 Hz，指令 8000 Hz 被钳位并置 0003_0131，
 *      波形一高一低各一拍；
 *   V3 限位：正向运动中 bLimitPos → 本拍停发、锁 0003_02E1、报警字 bit0；
 *      复位后仍拒正向（0003_0134），反向受理；
 *   V4 堵转：理论 1 s、裕度 500 ms → 2 s 到期锁 0003_02E3 并停发；
 *   V5 停车：运动中 Stop → 剩余步数压到减速段，频率降零回空闲，位置与已发
 *      脉冲数一致；
 *   V6 去使能：Enable(FALSE) → 本拍停发（无半脉冲）、bEnableOut FALSE、位置
 *      保持，再使能不自动续走。
 * 修订历史 (Revision)   :
 *   2026-11-15  v1.0.0  首版入库（Round 09 · DL_Device 开环步进族 · 实现件）
 *   2026-11-15  v1.0.1  终审修复：eDecel 补「频率归零即收尾」第二出口（原实现
 *                       仅在步数 <= 1E-6 时出口，减速段一拍归零而残差为小数时
 *                       状态机永久停在 eDecel，属无故障码的静默卡死）；新增
 *                       信息级 0003_0137 记录该收尾口径
 *============================================================================*)

(*-----------------------------------------------------------------------------
 * 调用示例 (Instance guide)：
 *   stCfg.uStepsPerMm := 400; stCfg.uMicrostep := 8; stCfg.fMaxSpeed := 30.0;
 *   stCfg.fAccel := 400.0; stCfg.tStallTimeout := T#300MS; stCfg.fTaskCycle := 0.01;
 *   bOk := fbStep.Init(stCfg := stCfg);      // 注入组态（调用方持有结构体）
 *   bOk := fbStep.Enable(bEnable := TRUE);   // 上使能（保持力矩）
 *   fbStep(bLimitPos := bDiPos, bLimitNeg := bDiNeg, bAlarmIn := bDiAlm);
 *   bOk := fbStep.MoveRelative(fDistance := 25.0, fSpeed := 15.0);
 *   上层映射：bDoPulse := fbStep.bPulse; bDoDir := fbStep.bDir;
 *   常见误用：① 脉宽硬下限——10 ms 任务最高 50 Hz，更高频率必须换更快的任务；
 *   ② 开环会丢步，fPosition 禁止当反馈做闭环；③ 有效当量 = 当量 × 细分，
 *   改细分必须同步改字段，否则速度与行程成比例偏差；④ 堵转判据识别卡滞不识别
 *   打滑；⑤ 故障期保持使能是有意设计（垂直轴防溜车），切动力请在安全回路侧。
 *----------------------------------------------------------------------------*)

(*-----------------------------------------------------------------------------
 * 枚举: E_DL_StepperState（归属 FB_DL_PulseDirStepper，随本文件发布）
 *----------------------------------------------------------------------------*)
{attribute 'strict'}
{attribute 'qualified_only'}
TYPE E_DL_StepperState :
(
    eIdle  := 0,     // 空闲待机：无运动，脉冲停发，可受理新指令 / Idle, pulses stopped and ready for a new command
    eAccel := 10,    // 加速段：频率按加速度斜坡上升 / Acceleration segment, frequency ramps up
    eRun   := 20,    // 匀速段：频率保持峰值 / Constant segment, frequency held at the peak
    eDecel := 30,    // 减速段：频率按减速度斜坡下降 / Deceleration segment, frequency ramps down
    eFault := 99     // 故障锁存：脉冲停发，仅复位可退 / Fault latched, only reset can leave
) UINT;
END_TYPE

FUNCTION_BLOCK FB_DL_PulseDirStepper IMPLEMENTS I_DL_StepperOpenLoop
VAR_INPUT
    bLimitPos    : BOOL;                // 正限位开关输入（Positive limit switch），TRUE = 触发；常闭型由调用方反相 / TRUE means triggered
    bLimitNeg    : BOOL;                // 负限位开关输入（Negative limit switch），TRUE = 触发 / TRUE means triggered
    bAlarmIn     : BOOL;                // 驱动器报警输入（Drive alarm input），TRUE = 报警 / TRUE means the drive reports an alarm
    fJogSpeed    : LREAL := 5.0;        // 点动速度预留（Reserved jog speed）[mm/s]，本版不启用 / Reserved, unused in this version
END_VAR
VAR_OUTPUT
    bPulse       : BOOL;                // 脉冲输出（Pulse output），定宽一拍（R24）/ Fixed one-scan-wide pulse per R24
    bDir         : BOOL;                // 方向输出（Direction output），TRUE = 正向 / TRUE means the positive direction
    bEnableOut   : BOOL;                // 使能输出（Enable output），透传指令，故障期保持 / Pass-through, held during faults
    fFreqNow     : LREAL;               // 当前脉冲频率（Current pulse frequency）[Hz]，诊断用 / Diagnostic frequency in hertz
    bError       : BOOL;                // 故障保持型（Fault latched），排除信息级码 / Latched fault flag, info codes excluded
    uErrorId     : UDINT;               // 故障码（Error code），0 = 无故障，段位 16#0003_xxxx / Error code, zero means no error
END_VAR
VAR
    _stCfg       : ST_DL_StepperCfg;    // 组态副本（Configuration copy），Init 注入 / Copy injected by Init
    _eState      : E_DL_StepperState := E_DL_StepperState.eIdle; // 主状态机状态（Main state machine state）/ Main state machine state
    _bInit       : BOOL;                // 首扫完成标志（First-scan done flag），初值 FALSE / First-scan done flag, initial FALSE
    _bInited     : BOOL;                // 组态已注入标志（Configuration injected flag）/ Configuration injected flag
    _bEnableCmd  : BOOL;                // 使能指令电平（Enable command level），Enable 方法写入 / Written by the Enable method
    _bPendMove   : BOOL;                // 待受理运动请求（Pending move request），方法置位主体消化 / Set by the method, consumed by the body
    _bPendStop   : BOOL;                // 待受理停车请求（Pending stop request），方法置位主体消化 / Set by the method, consumed by the body
    _bPendReset  : BOOL;                // 待受理复位请求（Pending reset request），方法置位主体消化 / Set by the method, consumed by the body
    _fPendDist   : LREAL;               // 待受理位移（Pending distance）[mm]，带符号 / Signed pending distance [mm]
    _fPendSpeed  : LREAL;               // 待受理速度（Pending speed）[mm/s]，已钳位 / Clamped pending speed [mm/s]
    _fPulsePerMm : LREAL := 400.0;      // 有效脉冲当量（Effective pulses per millimetre）[脉冲/mm]=当量×细分 / Equivalent times microstep divisor
    _fTaskCycle  : LREAL := 0.01;       // 生效任务周期（Effective task cycle）[s] / Effective task cycle [s]
    _fFreqMaxScan : LREAL := 50.0;      // 周期决定的频率上限（Cycle-driven frequency limit）[Hz]=1/(2×周期) / One over twice the cycle
    _fAccStepHz  : LREAL := 200000.0;   // 脉冲域加速度（Acceleration in the pulse domain）[脉冲/s²]=加速度×当量 / Acceleration scaled to pulses
    _fFreqStepHz : LREAL := 2000.0;     // 每拍频率增量（Frequency step per scan）[Hz]=脉冲域加速度×周期 / Pulse acceleration times the cycle
    _fFreqCmd    : LREAL;               // 指令频率（Command frequency）[Hz]，钳位后 / Command frequency after clamping [Hz]
    _fFreqTarget : LREAL;               // 峰值频率（Peak frequency）[Hz]，梯形峰值 / Trapezoidal peak frequency [Hz]
    _fFreqNow    : LREAL;               // 当前频率（Current frequency）[Hz]，逐拍积分 / Integrated frequency of this scan [Hz]
    _fStepsTotal : LREAL;               // 本次总步数（Total steps of this move）[脉冲]，正数 / Total pulses, always positive
    _fStepsRemain: LREAL;               // 剩余步数（Remaining steps）[脉冲]，递减到零即到位 / Counted down to zero on completion
    _fStepsAccel : LREAL;               // 加速段步数（Acceleration steps）[脉冲] / Pulses spent accelerating
    _fStepsDecel : LREAL;               // 减速段步数（Deceleration steps）[脉冲]，与加速段对称 / Symmetric with the acceleration segment
    _fPhaseAcc   : LREAL;               // 脉冲相位累加器（Pulse phase accumulator）[周期]，域 0 至 1 / Phase accumulator, zero to one period
    _fPosSteps   : LREAL;               // 指令位置脉冲数（Command position in pulses）[脉冲]，带符号 / Signed accumulated command position
    _fPosMm      : LREAL;               // 指令位置（Command position）[mm]，开环推算 / Open-loop derived command position [mm]
    _fExpectSec  : LREAL;               // 理论运动耗时（Theoretical move time）[s] / Theoretical move time [s]
    _fLimitSec   : LREAL;               // 堵转判据时限（Stall limit time）[s] / Stall limit time [s]
    _tMoveLimit  : TIME;                // 堵转判据时限（Stall limit as TIME）[ms]，喂定时器 / Stall limit fed to the timer [ms]
    _bMoveActive : BOOL;                // 运动进行中（Move active flag）/ Move active flag
    _bMoveBreak  : BOOL;                // 定时器断输入一拍（Timer break），运动起点重计时（公约 0.6）/ One-scan break at the move start
    _bDirNow     : BOOL;                // 当前运动方向（Current move direction），TRUE = 正向 / TRUE means positive
    _bLimitIntr  : BOOL;                // 同向限位入侵（Same-direction limit intrusion）/ Intrusion in the running direction
    _bFaultLatch : BOOL;                // 故障锁存（Fault latch），仅复位路径清除 / Fault latch, cleared only by the reset path
    _bStallLat   : BOOL;                // 堵转锁存（Stall latched），供报警字 bit3 / Stall latch feeding alarm bit three
    _uErrInt     : UDINT;               // 故障级码寄存（Fault-level code register），锁存型 / Latched fault-level code register
    _uInfoCode   : UDINT;               // 本拍信息级码（Info code this scan），每拍重算 / Info code recomputed every scan
    _uInfoHold   : UDINT;               // 方法拍信息级码保持（Method info code hold），供下一拍主体透出 / Held one scan for the body to expose
    _uAlarmWord  : WORD;                // 报警字（Alarm word），bit0 至 bit3 有效 / Alarm word with bits zero to three used
    _fbMoveTimer : TON;                 // 运动耗时监控定时器（Move elapsed timer），无条件刷新 / Refreshed unconditionally every scan
END_VAR
VAR CONSTANT
    DL_FLOAT_EPS     : LREAL := 1.0E-6; // 浮点容差（Float epsilon）[mm]，替代判等 / Float epsilon replacing equality [mm]
    DL_FREQ_EPS      : LREAL := 0.1;    // 频率容差（Frequency epsilon）[Hz] / Frequency epsilon [Hz]
    DL_TIMEOUT_GAIN  : LREAL := 1.5;    // 堵转裕度系数（Stall timeout gain），理论耗时倍数 / Multiplier on the theoretical time
    DL_PHASE_FULL    : LREAL := 1.0;    // 相位满量程（Full phase period）[周期] / Full phase period in cycles
    DL_PHASE_GUARD   : LREAL := 1.5;    // 相位防越界上限（Phase guard bound）[周期] / Defensive phase clamp bound
    DL_CYCLE_FALLBACK : LREAL := 0.01;  // 任务周期兜底（Task cycle fallback）[s] / Fallback task cycle [s]
    DL_LIMIT_SEC_MAX : LREAL := 3600.0; // 时限上限（Upper bound of the limit）[s]，防溢出 / Bound preventing overflow [s]
    DL_ALM_LIMIT_POS : WORD := 16#0001; // 报警字 bit0 正限位（Alarm bit zero, positive limit）/ Positive limit alarm bit
    DL_ALM_LIMIT_NEG : WORD := 16#0002; // 报警字 bit1 负限位（Alarm bit one, negative limit）/ Negative limit alarm bit
    DL_ALM_DRIVE     : WORD := 16#0004; // 报警字 bit2 驱动器报警（Alarm bit two, drive alarm）/ Drive alarm bit
    DL_ALM_STALL     : WORD := 16#0008; // 报警字 bit3 堵转超时（Alarm bit three, stall timeout）/ Stall timeout alarm bit
END_VAR

METHOD Init : BOOL
VAR_IN_OUT
    stCfg : ST_DL_StepperCfg;          // 步进组态（Stepper configuration），调用方持有 / Caller-owned configuration
END_VAR
IF (stCfg.uStepsPerMm = 0) OR (stCfg.uMicrostep = 0) OR (stCfg.fMaxSpeed <= DL_FLOAT_EPS) OR
   (stCfg.fAccel <= DL_FLOAT_EPS) OR (stCfg.fTaskCycle <= DL_FLOAT_EPS) OR
   (stCfg.fMaxSpeed <> stCfg.fMaxSpeed) OR (stCfg.fAccel <> stCfg.fAccel) OR
   (stCfg.fTaskCycle <> stCfg.fTaskCycle) THEN
    _uErrInt     := 16#0003_02E0;      // 0003_02E0 组态参数非法【故障级】（Illegal configuration, fault level）
    _bFaultLatch := TRUE;              // 越界锁故障（Violation latches a fault）
    _bInited     := FALSE;             // 保持未初始化（Remains uninitialized）
    Init         := FALSE;             // 受理失败（Rejected）
ELSE
    _stCfg       := stCfg;             // 保存组态副本（Keep a copy）
    _bInited     := TRUE;              // 置已初始化（Mark initialized）
    _uErrInt     := 16#0000_0000;      // 故障码清零（Fault code cleared）
    _bFaultLatch := FALSE;             // 成功初始化解除参数锁存（Successful init releases the latch）
    Init         := TRUE;              // 受理成功（Accepted）
END_IF

// 方法: Enable —— 电平语义，TRUE 使能（故障态拒绝），FALSE 恒受理并冻结（Method Enable）
    END_METHOD

METHOD Enable : BOOL
VAR_INPUT
    bEnable : BOOL;                    // 使能指令（Enable command），TRUE = 使能 / TRUE enables
END_VAR
IF bEnable THEN
    IF (NOT _bInited) OR _bFaultLatch OR (_eState = E_DL_StepperState.eFault) THEN
        _uInfoHold := 16#0003_0133;    // 0003_0133 指令被拒绝【信息级】（Command rejected, info level）
        Enable     := FALSE;           // 未初始化或故障态拒绝（Refused while uninitialized or faulty）
    ELSE
        _bEnableCmd := TRUE;           // 登记使能（Enable registered）
        Enable      := TRUE;           // 受理成功（Accepted）
    END_IF
ELSE
    _bEnableCmd := FALSE;              // 去使能恒受理（Disable always accepted）
    Enable      := TRUE;               // 受理成功（Accepted）
END_IF

// 方法: MoveRelative —— 仅空闲态受理，参数与限位方向先行校验（Method MoveRelative）
    END_METHOD

METHOD MoveRelative : BOOL
VAR_INPUT
    fDistance : LREAL;                 // 相对位移（Relative distance）[mm]，带符号 / Signed distance [mm]
    fSpeed    : LREAL;                 // 运行速度（Run speed）[mm/s]，必需为正 / Must be positive
END_VAR
IF (NOT _bInited) OR (NOT _bEnableCmd) OR _bFaultLatch OR (_eState <> E_DL_StepperState.eIdle) OR
   (fDistance <> fDistance) OR (ABS(fDistance) <= DL_FLOAT_EPS) OR
   (fSpeed <> fSpeed) OR (fSpeed <= DL_FLOAT_EPS) THEN
    _uInfoHold   := 16#0003_0133;      // 0003_0133 指令被拒绝【信息级】（Command rejected, info level）
    MoveRelative := FALSE;             // 拒绝受理（Rejected）
ELSIF (fDistance > 0.0) AND bLimitPos THEN
    _uInfoHold   := 16#0003_0134;      // 0003_0134 限位方向禁止【信息级】（Direction blocked, info level）
    MoveRelative := FALSE;             // 正限位上禁止正向（Positive motion refused at the positive limit）
ELSIF (fDistance < 0.0) AND bLimitNeg THEN
    _uInfoHold   := 16#0003_0134;      // 0003_0134 限位方向禁止【信息级】（Direction blocked, info level）
    MoveRelative := FALSE;             // 负限位上禁止负向（Negative motion refused at the negative limit）
ELSE
    IF (_stCfg.fMaxSpeed > DL_FLOAT_EPS) AND (fSpeed > _stCfg.fMaxSpeed) THEN
        _fPendSpeed := _stCfg.fMaxSpeed; // 钳位到最大速度（Clamped to the maximum）
        _uInfoHold  := 16#0003_0130;     // 0003_0130 速度超限已钳位【信息级】（Speed clamped, info level）
    ELSE
        _fPendSpeed := fSpeed;          // 合法速度直通（Valid speed passed through）
    END_IF
    _fPendDist   := fDistance;          // 登记位移（Distance registered）
    _bPendMove   := TRUE;               // 登记运动请求（Move request registered）
    MoveRelative := TRUE;               // 受理成功（Accepted）
END_IF

// 方法: Stop —— 受控停车：剩余步数压到减速段后按斜坡降频（Method Stop）
    END_METHOD

METHOD Stop : BOOL
VAR_INPUT
END_VAR
IF _bMoveActive THEN
    _bPendStop := TRUE;                // 登记停车请求（Stop request registered）
    Stop       := TRUE;                // 受理成功（Accepted）
ELSE
    _uInfoHold := 16#0003_0133;        // 0003_0133 指令被拒绝【信息级】（Command rejected, info level）
    Stop       := FALSE;               // 无运动可停（Nothing to stop）
END_IF

// 方法: Reset —— 仅故障锁存时受理；报警源未消失则保留锁存（Method Reset）
    END_METHOD

METHOD Reset : BOOL
VAR_INPUT
END_VAR
IF _bFaultLatch OR (_eState = E_DL_StepperState.eFault) THEN
    _bPendReset := TRUE;               // 登记复位请求，主体按报警源裁决（Reset registered, body decides）
    Reset       := TRUE;               // 受理成功（Accepted）
ELSE
    _uInfoHold  := 16#0003_0133;       // 0003_0133 无故障可复位【信息级】（Nothing to reset, info level）
    Reset       := FALSE;              // 拒绝受理（Rejected）
END_IF

// 方法: GetErrorId —— 故障码查询，与 uErrorId 引脚同源（Method GetErrorId）
    END_METHOD

METHOD GetErrorId : UDINT
VAR_INPUT
END_VAR
GetErrorId := uErrorId;                // 直接透出末次码（Expose the last code）

// 属性: bReady（GET）—— 已初始化 + 已使能 + 无故障 + 空闲（Property bReady）
    END_METHOD

// 段 1｜出口确定性与单拍标志预清零（公约 0.9 / R25 第一律：停发在本拍内完成）
bPulse     := FALSE;                   // 脉冲默认低电平（Pulse defaults low）
_uInfoCode := _uInfoHold;              // 先透出方法拍产生的信息级码，保留单拍（Method codes survive one body scan）
_uInfoHold := 0;                       // 单拍消费后自清（Consumed and cleared after exactly one scan）
_bLimitIntr := FALSE;                  // 限位入侵标志每拍重算（Intrusion recomputed every scan）

// 段 2｜首扫初始化（R19 范式：IF (NOT _bInit) 唯一判据）
IF NOT _bInit THEN
    _bInit        := TRUE;             // 置首扫完成（First-scan done）
    _eState       := E_DL_StepperState.eIdle; // 状态复位空闲（State reset to idle）
    _bEnableCmd   := FALSE;            // 使能指令清零（Enable command cleared）
    _bPendMove    := FALSE;            // 清待受理运动（Pending move cleared）
    _bPendStop    := FALSE;            // 清待受理停车（Pending stop cleared）
    _bPendReset   := FALSE;            // 清待受理复位（Pending reset cleared）
    _fFreqNow     := 0.0;              // 当前频率清零（Frequency cleared）
    _fPhaseAcc    := 0.0;              // 相位累加器清零（Phase cleared）
    _fPosSteps    := 0.0;              // 位置脉冲数清零（Position pulses cleared）
    _fPosMm       := 0.0;              // 位置清零（Position cleared）
    _bMoveActive  := FALSE;            // 运动标志清零（Move flag cleared）
    _bDirNow      := TRUE;             // 方向默认正向（Direction defaults positive）
    _bFaultLatch  := FALSE;            // 故障锁存清零（Fault latch cleared）
    _bStallLat    := FALSE;            // 堵转锁存清零（Stall latch cleared）
    _uErrInt      := 16#0000_0000;     // 故障码清零（Fault code cleared）
    _uAlarmWord   := 16#0000;          // 报警字清零（Alarm word cleared）
END_IF

// 段 3｜定时器无条件刷新（公约 0.5 / 0.6：断输入一拍后从零重计）
_fbMoveTimer(IN := _bMoveActive AND (NOT _bMoveBreak), PT := _tMoveLimit); // 运动耗时监控（Move elapsed monitoring）
_bMoveBreak := FALSE;                  // 断输入脉冲在实例调用后自清（Break self-cleared after the call）

// 段 4｜组态派生与参数防御（脉冲域换算、频率上限、除零守卫）
IF _bInited THEN
    IF (_stCfg.fTaskCycle <> _stCfg.fTaskCycle) OR (_stCfg.fTaskCycle <= DL_FLOAT_EPS) THEN
        _fTaskCycle := DL_CYCLE_FALLBACK; // 周期非法兜底（Illegal cycle falls back）
        _uInfoCode  := 16#0003_0136;      // 0003_0136 任务周期非法已兜底【信息级】（Cycle fell back, info level）
    ELSE
        _fTaskCycle := _stCfg.fTaskCycle; // 合法周期直通（Valid cycle passed through）
    END_IF
    _fPulsePerMm := UINT_TO_LREAL(_stCfg.uStepsPerMm) * UINT_TO_LREAL(_stCfg.uMicrostep); // 有效当量（Effective equivalent）
    IF _fPulsePerMm <= DL_FLOAT_EPS THEN
        _bFaultLatch := TRUE;          // 当量为零锁故障（Zero equivalent latches a fault）
        _uErrInt     := 16#0003_02E0;  // 0003_02E0 组态参数非法【故障级】（Illegal configuration, fault level）
        _fPulsePerMm := 1.0;           // 除零守卫置 1（Divide guard set to one）
    END_IF
    _fFreqMaxScan := 1.0 / (2.0 * _fTaskCycle); // 频率上限，脉宽下限一拍（Ceiling keeping the pulse one scan wide）
    _fAccStepHz   := _stCfg.fAccel * _fPulsePerMm; // 脉冲域加速度 [脉冲/s²]（Pulse-domain acceleration）
    _fFreqStepHz  := _fAccStepHz * _fTaskCycle;    // 每拍频率增量 [Hz]（Frequency increment per scan）
END_IF

// 段 5｜故障源监视与锁存（限位入侵 / 驱动器报警 / 堵转超时；0.7 锁存型）
_bLimitIntr := _bMoveActive AND ((_bDirNow AND bLimitPos) OR ((NOT _bDirNow) AND bLimitNeg)); // 同向限位判据（Intrusion verdict）
IF _bMoveActive THEN
    IF _bLimitIntr THEN
        _bFaultLatch := TRUE;          // 限位入侵锁存（Intrusion latched）
        _uErrInt     := 16#0003_02E1;  // 0003_02E1 限位入侵停机【故障级】（Intrusion stop, fault level）
    ELSIF bAlarmIn THEN
        _bFaultLatch := TRUE;          // 驱动器报警锁存（Drive alarm latched）
        _uErrInt     := 16#0003_02E2;  // 0003_02E2 驱动器报警输入【故障级】（Drive alarm, fault level）
    ELSIF _fbMoveTimer.Q THEN
        _bFaultLatch := TRUE;          // 堵转超时锁存（Stall timeout latched）
        _bStallLat   := TRUE;          // 报警字 bit3 保持（Alarm bit three held）
        _uErrInt     := 16#0003_02E3;  // 0003_02E3 堵转超时【故障级】（Stall timeout, fault level）
    END_IF
END_IF

// 段 6｜请求消化：复位（报警源优先）/ 停车（受控减速）/ 去使能（本拍冻结）
IF _bPendReset THEN
    _bPendReset := FALSE;              // 复位请求单拍消费（Reset request consumed）
    IF NOT bAlarmIn THEN
        _bFaultLatch := FALSE;         // 报警源消失才解除（Cleared only when the alarm is gone）
        _bStallLat   := FALSE;         // 堵转锁存解除（Stall latch released）
        _uErrInt     := 16#0000_0000;  // 故障码清零（Fault code cleared）
        IF _eState = E_DL_StepperState.eFault THEN
            _eState := E_DL_StepperState.eIdle; // 故障态退回空闲（Fault returns to idle）
        END_IF
    END_IF
END_IF
IF _bPendStop THEN
    _bPendStop := FALSE;               // 停车请求单拍消费（Stop request consumed）
    IF (_eState = E_DL_StepperState.eAccel) OR (_eState = E_DL_StepperState.eRun) THEN
        IF _fStepsRemain > _fStepsDecel THEN
            _fStepsRemain := _fStepsDecel; // 剩余步数压到减速段长度（Cut to the deceleration length）
        END_IF
        _eState := E_DL_StepperState.eDecel; // 进减速段受控停车（Controlled stop via deceleration）
    END_IF
END_IF
IF NOT _bEnableCmd THEN
    IF _bMoveActive THEN
        _uInfoCode := 16#0003_0135;    // 0003_0135 去使能冻结脉冲输出【信息级】（Disable freezes pulses, info level）
    END_IF
    _eState      := E_DL_StepperState.eIdle; // 去使能立即回空闲（Disable returns to idle）
    _fFreqNow    := 0.0;               // 频率清零（Frequency cleared）
    _fPhaseAcc   := 0.0;               // 相位清零，杜绝半脉冲（Phase cleared, no half pulse remains）
    _bMoveActive := FALSE;             // 运动标志清零（Move flag cleared）
    _fStepsRemain := 0.0;              // 剩余步数清零（Remaining steps cleared）
END_IF

// 段 7｜主状态机与梯形频率规划（ENUM + CASE + ELSE 兜底）
CASE _eState OF
    E_DL_StepperState.eIdle: // 空闲：等待运动请求（Idle, waiting for a move request）
        _fFreqNow    := 0.0;       // 空闲频率为零（Idle frequency is zero）
        _bMoveActive := FALSE;     // 空闲无运动（No motion while idle）
        IF _bFaultLatch THEN
            _eState := E_DL_StepperState.eFault; // 故障优先（Fault takes priority）
        ELSIF _bPendMove THEN
            _bPendMove := FALSE;   // 运动请求单拍消费（Move request consumed）
            _fStepsTotal := ABS(_fPendDist) * _fPulsePerMm; // 总步数 [脉冲]（Total pulses）
            IF _fStepsTotal <= DL_FLOAT_EPS THEN
                _uInfoCode := 16#0003_0132; // 0003_0132 位移不足一当量【信息级】（Distance below one pulse, info level）
            ELSE
                _fFreqCmd := _fPendSpeed * _fPulsePerMm; // 指令频率 [Hz]（Command frequency）
                IF _fFreqCmd > _fFreqMaxScan THEN
                    _fFreqCmd  := _fFreqMaxScan;         // 钳位到周期上限（Clamp to the cycle ceiling）
                    _uInfoCode := 16#0003_0131;          // 0003_0131 频率超上限已钳位【信息级】（Clamped, info level）
                END_IF
                IF _fAccStepHz > DL_FLOAT_EPS THEN
                    _fStepsAccel := (_fFreqCmd * _fFreqCmd) / (2.0 * _fAccStepHz); // na = v²/(2a)（Acceleration pulses）
                ELSE
                    _fStepsAccel := 0.0;                     // 加速度为零无加速段（No acceleration segment）
                END_IF
                IF (2.0 * _fStepsAccel) > _fStepsTotal THEN
                    _fStepsAccel := _fStepsTotal / 2.0;      // 三角型取半程（Triangular, half of the travel）
                    IF _fAccStepHz > DL_FLOAT_EPS THEN
                        _fFreqTarget := SQRT(_fAccStepHz * _fStepsTotal); // 峰值 = SQRT(a×N)（Triangular peak）
                    ELSE
                        _fFreqTarget := _fFreqCmd;           // 无加速度退化匀速（Constant speed fallback）
                    END_IF
                    IF _fFreqTarget > _fFreqCmd THEN
                        _fFreqTarget := _fFreqCmd;           // 峰值不超指令频率（Peak never exceeds the command）
                    END_IF
                ELSE
                    _fFreqTarget := _fFreqCmd;               // 梯形峰值 = 指令频率（Trapezoidal peak）
                END_IF
                _fStepsDecel  := _fStepsAccel;               // 减速段对称（Symmetric deceleration）
                _fStepsRemain := _fStepsTotal;               // 剩余步数装载（Remaining steps loaded）
                _fPhaseAcc    := 0.0;                        // 相位从头开始（Phase restarts）
                _bDirNow      := (_fPendDist > 0.0);         // 方向取位移符号（Direction from the sign）
                _bMoveActive  := TRUE;                       // 置运动进行中（Move marked active）
                _bMoveBreak   := TRUE;                       // 定时器下拍从零重计（Timer restarts next scan）
                _fExpectSec   := 0.0;                        // 理论耗时先清零（Theoretical time cleared）
                IF (_fFreqTarget > DL_FREQ_EPS) AND (_fAccStepHz > DL_FLOAT_EPS) THEN
                    _fExpectSec := (2.0 * (_fFreqTarget / _fAccStepHz)) +
                                   ((_fStepsTotal - (2.0 * _fStepsAccel)) / _fFreqTarget); // t = 2(v/a)+(N−2na)/v（Theoretical time）
                END_IF
                _fLimitSec := (_fExpectSec * DL_TIMEOUT_GAIN) +
                              (UDINT_TO_LREAL(TIME_TO_UDINT(_stCfg.tStallTimeout)) / 1000.0); // 时限 = 理论×裕度 + 附加裕度（Limit with margin）
                _fLimitSec := LIMIT(0.001, _fLimitSec, DL_LIMIT_SEC_MAX);                     // 防 TIME 溢出（Bound preventing overflow）
                _tMoveLimit := UDINT_TO_TIME(LREAL_TO_UDINT(_fLimitSec * 1000.0));            // 毫秒量化（Whole milliseconds）
                _eState := E_DL_StepperState.eAccel;         // 进加速段（Enter acceleration）
            END_IF
        END_IF

    E_DL_StepperState.eAccel: // 加速段：频率斜坡上升（Frequency ramps up）
        _fFreqNow := _fFreqNow + _fFreqStepHz; // 每拍加一增量（Advance one frequency step）
        IF _fFreqNow >= _fFreqTarget THEN
            _fFreqNow := _fFreqTarget;     // 到峰值封顶（Clamped at the peak）
            _eState   := E_DL_StepperState.eRun; // 转匀速段（Go to constant speed）
        END_IF
        IF _fFreqNow <= DL_FREQ_EPS THEN
            _fFreqNow := DL_FREQ_EPS;      // 起步频率守卫，防相位不累加（Startup guard）
        END_IF
        IF _fStepsRemain <= _fStepsDecel THEN
            _eState := E_DL_StepperState.eDecel; // 剩余步入减速区（Deceleration zone reached）
        END_IF

    E_DL_StepperState.eRun: // 匀速段：频率保持峰值（Constant segment）
        _fFreqNow := _fFreqTarget;         // 频率恒定（Frequency held）
        IF _fStepsRemain <= _fStepsDecel THEN
            _eState := E_DL_StepperState.eDecel; // 进减速段（Enter deceleration）
        END_IF

    E_DL_StepperState.eDecel: // 减速段：频率斜坡下降（Frequency ramps down）
        _fFreqNow := _fFreqNow - _fFreqStepHz; // 每拍减一增量（Retreat one frequency step）
        IF _fFreqNow <= DL_FREQ_EPS THEN
            _fFreqNow := 0.0;              // 频率归零（Frequency reaches zero）
        END_IF
        (* 收尾双出口（v1.0.1 终审补第二出口，状态终态可达性）：
           ① 步数走完 → 正常到位；
           ② 频率已归零 → 相位不再累加，剩余脉冲在数学上永不可发，必须按到位
              收尾；否则状态机永久停在 eDecel，表现为 bPulse 恒 FALSE、
              bError FALSE、bReady 恒 FALSE 的静默卡死。
              触发条件：每拍频率步进 fAccel×当量×周期 远大于峰值频率时
              （默认组态 2000 Hz/拍 vs 50 Hz 峰值即属此列），减速段一拍归零
              而残余分步（位移×当量带小数）尚未发完。 *)
        IF (_fStepsRemain <= DL_FLOAT_EPS) OR (_fFreqNow <= DL_FREQ_EPS) THEN
            IF _fStepsRemain > DL_FLOAT_EPS THEN
                _uInfoCode := 16#0003_0137; // 0003_0137 残差不足一脉冲按到位收尾【信息级】（Residual below one pulse, info level）
            END_IF
            _eState      := E_DL_StepperState.eIdle; // 步数归零回空闲（Idle when no step remains）
            _bMoveActive := FALSE;         // 运动结束（Move finished）
            _fFreqNow    := 0.0;           // 频率清零（Frequency cleared）
            _fPhaseAcc   := 0.0;           // 相位清零，杜绝残余半脉冲（Phase cleared, no half pulse remains）
        END_IF

    E_DL_StepperState.eFault: // 故障锁存：脉冲停发（Fault latched, pulses stopped）
        _fFreqNow     := 0.0;              // 频率清零（Frequency cleared）
        _bMoveActive  := FALSE;            // 运动标志清零（Move flag cleared）
        _fStepsRemain := 0.0;              // 剩余步数清零（Remaining steps cleared）

    ELSE
        _bFaultLatch := TRUE;              // 非法状态兜底锁存（Illegal state latched）
        _uErrInt     := 16#0003_02E4;      // 0003_02E4 非法状态兜底【故障级】（Illegal state, fault level）
        _eState      := E_DL_StepperState.eFault; // 进故障态（Enter the fault state）
        _fFreqNow    := 0.0;               // 频率清零（Frequency cleared）
        _bMoveActive := FALSE;             // 运动标志清零（Move flag cleared）
END_CASE

// 段 8｜脉冲发生（相位累加、定宽输出、步数与位置累计；R24 无半脉冲）
IF _bMoveActive AND (_fFreqNow > DL_FREQ_EPS) THEN
    _fPhaseAcc := _fPhaseAcc + (_fFreqNow * _fTaskCycle); // 相位增量 = 频率×周期（Phase increment）
    IF _fPhaseAcc > DL_PHASE_GUARD THEN
        _fPhaseAcc := DL_PHASE_FULL;   // 防御钳位，杜绝静默丢脉冲（Defensive clamp, no silent pulse loss）
    END_IF
    IF _fPhaseAcc >= DL_PHASE_FULL THEN
        _fPhaseAcc := _fPhaseAcc - DL_PHASE_FULL; // 消耗一个脉冲周期（Consume one period）
        bPulse := TRUE;                // 本拍输出一个定宽脉冲（Emit one fixed-width pulse）
        _fStepsRemain := _fStepsRemain - 1.0; // 剩余步数递减（Remaining steps decremented）
        IF _bDirNow THEN
            _fPosSteps := _fPosSteps + 1.0; // 正向累计（Accumulate positive）
        ELSE
            _fPosSteps := _fPosSteps - 1.0; // 负向累计（Accumulate negative）
        END_IF
    END_IF
END_IF
IF _bMoveActive AND (_fStepsRemain <= DL_FLOAT_EPS) THEN
    _eState      := E_DL_StepperState.eIdle; // 步数走完回空闲（Idle once every step is emitted）
    _bMoveActive := FALSE;             // 运动结束（Move finished）
    _fFreqNow    := 0.0;               // 频率清零（Frequency cleared）
    _fPhaseAcc   := 0.0;               // 相位清零（Phase cleared）
END_IF

// 段 9｜出口映射（位置、报警字、故障级码优先透出）
IF _fPulsePerMm > DL_FLOAT_EPS THEN
    _fPosMm := _fPosSteps / _fPulsePerMm; // 位置换算 [mm]（Position conversion）
ELSE
    _fPosMm := 0.0;                    // 除零守卫，位置报零（Divide guard, position reported as zero）
END_IF
bDir       := _bDirNow;                // 方向输出（Direction output）
bEnableOut := _bEnableCmd;             // 使能透传，故障期保持力矩（Enable passed through for holding torque）
fFreqNow   := _fFreqNow;               // 当前频率出口（Current frequency outlet）
_uAlarmWord := 16#0000;                // 报警字先清零（Alarm word cleared first）
IF bLimitPos THEN
    _uAlarmWord := _uAlarmWord OR DL_ALM_LIMIT_POS; // bit0 正限位（Positive limit bit）
END_IF
IF bLimitNeg THEN
    _uAlarmWord := _uAlarmWord OR DL_ALM_LIMIT_NEG; // bit1 负限位（Negative limit bit）
END_IF
IF bAlarmIn THEN
    _uAlarmWord := _uAlarmWord OR DL_ALM_DRIVE;     // bit2 驱动器报警（Drive alarm bit）
END_IF
IF _bStallLat THEN
    _uAlarmWord := _uAlarmWord OR DL_ALM_STALL;     // bit3 堵转超时保持（Stall timeout bit, held）
END_IF
bError := _bFaultLatch OR (_eState = E_DL_StepperState.eFault); // 故障派生，排除信息级（Fault derived, info codes excluded）
IF bError THEN
    uErrorId := _uErrInt;              // 故障级码优先（Fault-level code first）
ELSE
    uErrorId := _uInfoCode;            // 无故障透出信息级码（Info code exposed）
END_IF

// 方法: Init —— 注入组态并校验参数域，越界锁故障（Method Init, configuration validation）

PROPERTY bReady : BOOL
bReady := _bInited AND _bEnableCmd AND (NOT _bFaultLatch) AND (_eState = E_DL_StepperState.eIdle); // 就绪派生式（Ready derived form）

// 属性: fPosition（GET）—— 指令位置累计，开环推算非反馈（Property fPosition）
PROPERTY fPosition : LREAL
fPosition := _fPosMm;                  // 透出内部位置（Expose the internal position）

// 属性: uAlarmWord（GET）—— 报警字位域回读（Property uAlarmWord）
PROPERTY uAlarmWord : WORD
uAlarmWord := _uAlarmWord;             // 透出内部报警字（Expose the internal alarm word）
END_FUNCTION_BLOCK
